Staubli VAL3: insertAction.pgx

public program insertAction()
  local bool l_bExit
  local num l_i
  local num l_nActionIndex
  local bool l_bResult
  local num l_nPoint
  local bool l_bResult1
begin
  do
    if util:sPage!="insertAction"
      util:sPage="insertAction"
      resize(sActionList,1,size(actiondata:aActItem))
      for l_i = 0 to size(sActionList)-1
        sActionList[l_i]=toString("",l_i)+","+actiondata:aActItem[l_i].sComment
      endFor
      sSelAction=""
      userPageBind("insertAction","cbx1","options",sActionList,size(sActionList),"r")
      userPageBind("insertAction","cbx1","value",sSelAction,1,"rw")
      userPageBindClick("insertAction","btn1",bAConfirm,true)
      userPageBindClick("insertAction","btn2",bACancel,true)
      userPage(util:sPage)
      delay(0.5)
    endIf
    //
    if bAConfirm
      bAConfirm=false
      call trajectory:getPointIndex(sTrajItem,sSelPoint,l_nPoint,l_bResult1)
      toNum(sSelAction,l_nActionIndex,l_bResult)
      if l_bResult
        call trajectory:insertAction(sTrajItem,l_nPoint,l_nActionIndex,bToSave)
        l_bExit=true
      else
        userPageAlert("选择正确的action")
      endIf
    elseIf bACancel
      bACancel=false
      l_bExit=true

    endIf

    delay(0)
  until l_bExit==true
end
